TYPE ST_MotionFunctionPoint :
STRUCT
	nPointIndex: UDINT;
	nNextPointIndex: UDINT;
	eFunctionType: E_MotionFunctionType;
	ePointType: E_MotionPointType;
	/// X 
	MasterPos: LREAL;
	/// Y 
	SlavePos: LREAL;
	/// Y' 
	SlaveVelo: LREAL;
	/// Y'' 
	SlaveAcc: LREAL;
	/// Y''' 
	SlaveJerk: LREAL;
END_STRUCT
END_TYPE

(* stored: Version 1.1.0.1, ProductVersion 3.1.4024.12
   DUT ST_MotionFunctionPoint: Id {ebe2ed35-1f3a-4e00-b48d-8b9a5c5998f1} *)
